(* PLC project 未命名, 未知 未命名 1 *)
(* stored: creationDateTime 2025-05-30T09:25:40, modificationDateTime 2025-06-05T10:41:41 *)

PROGRAM program0
  VAR
    Up AT %IX0.1 : BOOL;
    Down AT %IX0.3 : BOOL;
    Start AT %IX0.6 : BOOL := 0;
    Stop AT %IX0.0 : BOOL := 0;
    Emergency AT %IX0.2 : BOOL;
    Working_LED AT %QX0.0 : BOOL;
    LED1 AT %QX0.1 : BOOL;
    LED2 AT %QX0.2 : BOOL;
    LED3 AT %QX0.3 : BOOL;
    LED4 AT %QX0.4 : BOOL;
    LED5 AT %QX0.5 : BOOL;
    LED6 AT %QX0.6 : BOOL;
  END_VAR
  VAR
    CTUD0 : CTUD;
    Run : BOOL;
    Run0 : BOOL;
    CV : INT := 5;
    CT : INT := 5;
  END_VAR
  VAR  (* added by the conversion: wires and edge detectors of the diagram *)
    R_TRIG1 : R_TRIG;
    R_TRIG2 : R_TRIG;
    _EQ49_OUT : BOOL;
    _EQ51_OUT : BOOL;
    _EQ53_OUT : BOOL;
    _EQ57_OUT : BOOL;
    _EQ56_OUT : BOOL;
    R_TRIG3 : R_TRIG;
  END_VAR

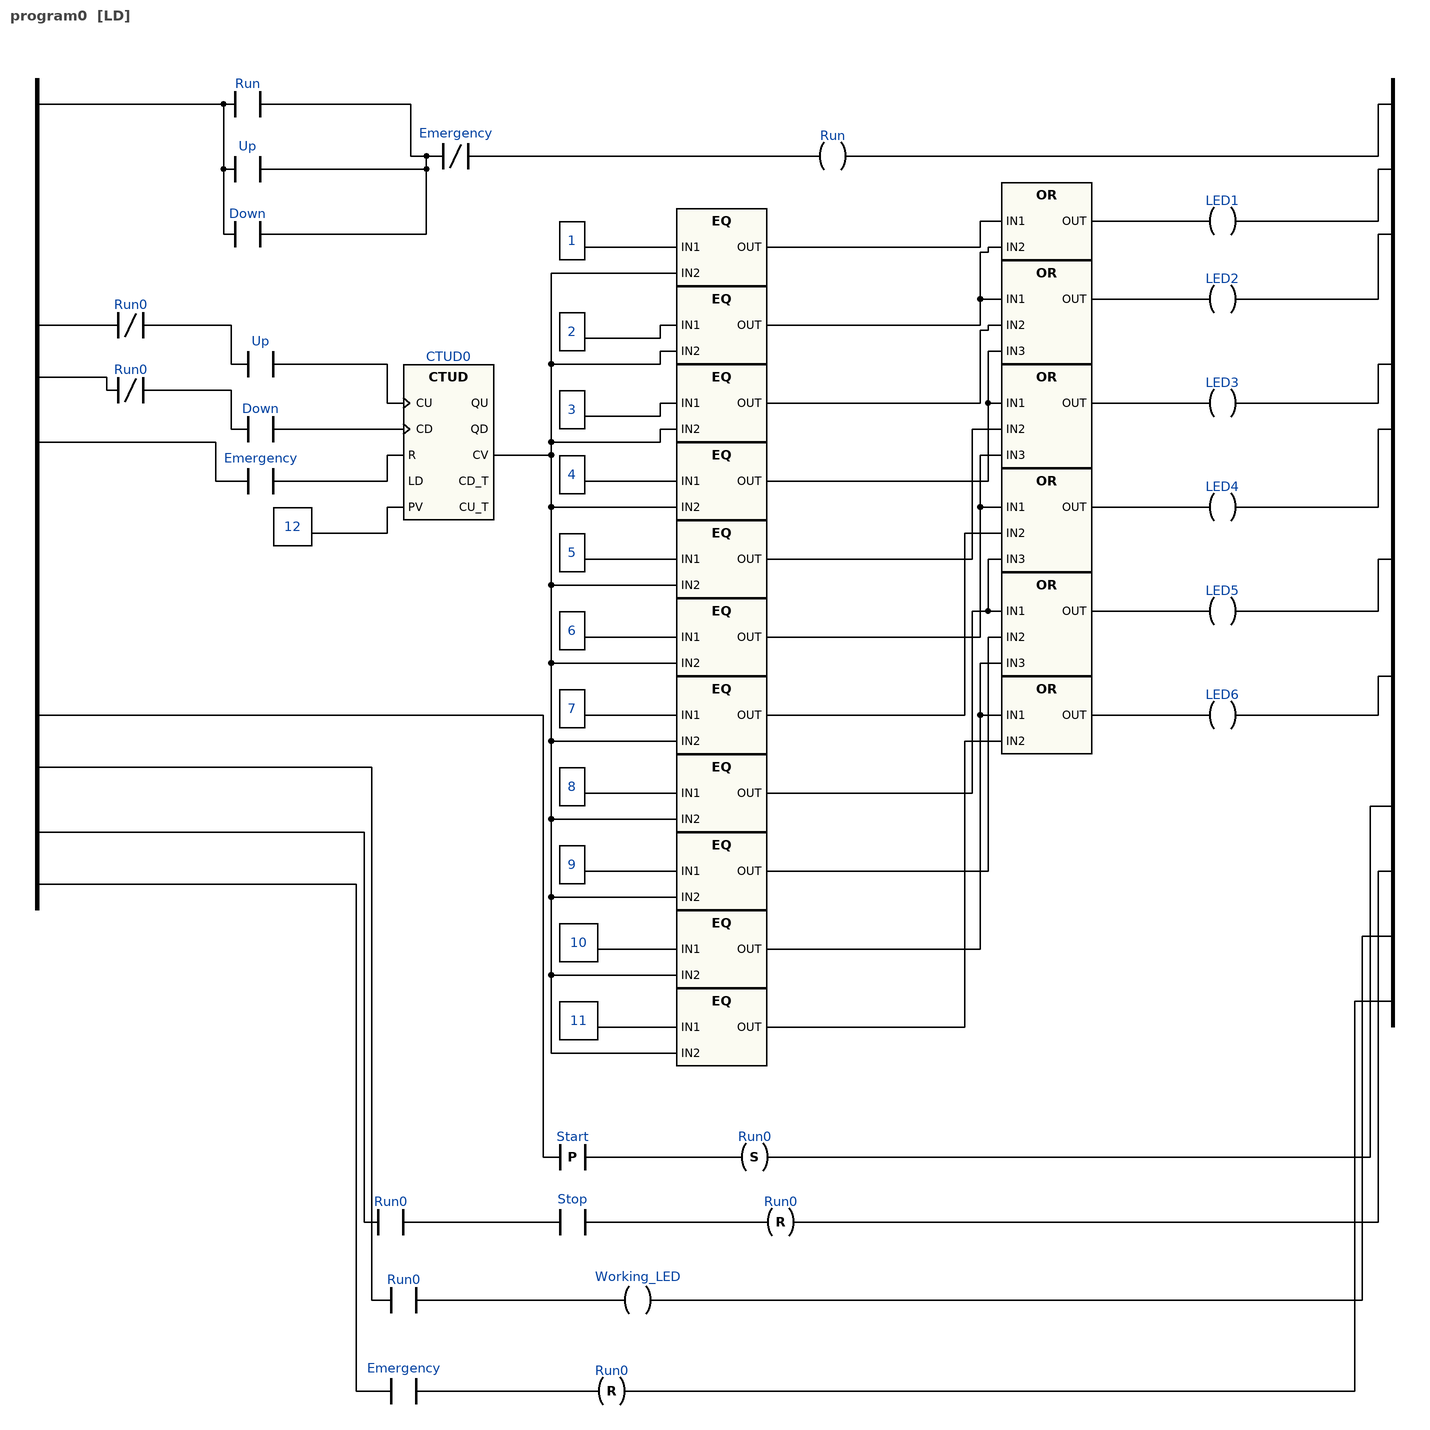
(* LD diagram, written out as Structured Text *)
Run := (Run OR Up OR Down) AND NOT Emergency;
R_TRIG1(CLK := NOT Run0 AND Up);
R_TRIG2(CLK := NOT Run0 AND Down);
CTUD0(CU := R_TRIG1.Q, CD := R_TRIG2.Q, R := Emergency, PV := 12);
_EQ49_OUT := 2 = CTUD0.CV;
LED1 := 1 = CTUD0.CV OR _EQ49_OUT;
_EQ51_OUT := 4 = CTUD0.CV;
LED2 := _EQ49_OUT OR 3 = CTUD0.CV OR _EQ51_OUT;
_EQ53_OUT := 6 = CTUD0.CV;
LED3 := _EQ51_OUT OR 5 = CTUD0.CV OR _EQ53_OUT;
_EQ57_OUT := 8 = CTUD0.CV;
LED4 := _EQ53_OUT OR 7 = CTUD0.CV OR _EQ57_OUT;
_EQ56_OUT := 10 = CTUD0.CV;
LED5 := _EQ57_OUT OR 9 = CTUD0.CV OR _EQ56_OUT;
LED6 := _EQ56_OUT OR 11 = CTUD0.CV;
IF Run0 AND Stop THEN Run0 := FALSE; END_IF;
R_TRIG3(CLK := Start);
IF R_TRIG3.Q THEN Run0 := TRUE; END_IF;
Working_LED := Run0;
IF Emergency THEN Run0 := FALSE; END_IF;
END_PROGRAM

CONFIGURATION Config0
  RESOURCE Res0 ON PLC
    TASK mytask(INTERVAL := T#100ms, PRIORITY := 1);
    PROGRAM mainLogic WITH mytask : program0;
  END_RESOURCE
END_CONFIGURATION
